Universal Robots URScript: TgtProg.script

def TgtProg():
  # Global parameters:
  global speed_ms    = 0.250
  global speed_rads  = 0.750
  global accel_mss   = 1.200
  global accel_radss = 1.200
  global blend_radius_m = 0.001
  global ref_frame = p[0,0,0,0,0,0]

  #
  # TO REMOVE HEADER:
  # Go to "Program" -> "Post-Processor Editor"
  # Select "Universal Robots"
  # Set "INCLUDE_HEADER" to "False"
  #
  #--------------------------
  # Add any default subprograms here
  # For example, to drive a gripper as a program call:
  # def Gripper_Open():
  #   ...
  # end
  #
  # Example to drive a spray gun:
  def SprayOn(value):
    # use the value as an output:
    DO_SPRAY = 5
    if value == 0:
      set_standard_digital_out(DO_SPRAY, False)
    else:
      set_standard_digital_out(DO_SPRAY, True)
    end
  end

  # Example to drive an extruder:
  def Extruder(value):
    # use the value as an output:
    if value < 0:
      # stop extruder
    else:
      # start extruder
    end
  end

  # Example to move an external axis
  def MoveAxis(value):
    # use the value as an output:
    DO_AXIS_1 = 1
    DI_AXIS_1 = 1
    if value <= 0:
      set_standard_digital_out(DO_AXIS_1, False)

      # Wait for digital input to change state
      #while (get_standard_digital_in(DI_AXIS_1) != False):
      #  sync()
      #end
    else:
      set_standard_digital_out(DO_AXIS_1, True)

      # Wait for digital input to change state
      #while (get_standard_digital_in(DI_AXIS_1) != True):
      #  sync()
      #end
    end
  end
  #--------------------------


  # Main program:
  # Program generated by RoboDK v6.0.7 for UR10 on XX/XX/XXXX 18:00:00
  # Using nominal kinematics.
  set_standard_digital_out(0, True)
  set_standard_digital_out(7, True)
  set_standard_digital_out(9, True)
  set_tool_digital_out(0, True)
  set_tool_digital_out(2, True)
  set_tool_digital_out(9, True)
  set_configurable_digital_out(0, True)
  set_configurable_digital_out(80, True)
  set_standard_digital_out(-1, True)
  set_standard_digital_out(1, False)
  set_standard_digital_out(1, True)
  set_standard_digital_out(1, False)
  set_standard_digital_out(1, True)
  set_standard_digital_out(1, False)
  set_standard_digital_out(1, False)
  set_standard_digital_out(1, True)
  set_standard_digital_out(1, True)
  set_standard_digital_out(1, true)
  set_standard_digital_out(1, TRUE)
  set_standard_digital_out(1, tRuE)
  set_standard_digital_out(1, False)
  set_standard_digital_out(1, False)
  set_standard_digital_out(1, False)
  A = B
  A = 1
  1 = 1
  # End of main program
end

TgtProg()
